(* IEC 61131-3 sources: engineering-notes/하드웨어코딩_hardware-coding/현업언어_industry-languages/04-PLC스캔_structured-text, 1 file *)

(* ---- indicator.st ---- *)
FUNCTION_BLOCK TempIndicator (* 호출 사이에 표시 상태를 기억할 블록 *)
VAR_INPUT (* 매 스캔에 전달할 입력 *)
    Enable : BOOL; (* 표시 기능의 사용 여부 *)
    Temperature10 : DINT; (* 온도 0.1도 단위의 정수 표본 *)
END_VAR (* 입력 선언 끝 *)
VAR_OUTPUT (* 호출 뒤 읽을 출력 *)
    Lit : BOOL := FALSE; (* 시작할 때 표시등은 꺼 두기 *)
END_VAR (* 출력 선언 끝 *)
IF NOT Enable THEN (* 사용하지 않으면 이전 상태보다 우선 *)
    Lit := FALSE; (* 표시 상태 지우기 *)
ELSIF Temperature10 >= 300 THEN (* 30.0도부터 켜기 *)
    Lit := TRUE; (* 높은 구간에서 켜진 상태 저장 *)
ELSIF Temperature10 <= 250 THEN (* 25.0도까지 내려오면 끄기 *)
    Lit := FALSE; (* 낮은 구간에서 꺼진 상태 저장 *)
END_IF; (* 중간 구간에서는 대입하지 않아 직전 상태 유지 *)
END_FUNCTION_BLOCK (* 한 번 호출이 한 번의 상태 갱신 *)
